(* IEC 61131-3 sources: iec-checker/test/st/bad, 2 files *)

(* ---- semantic-error.st ---- *)
TYPE
  ANALOG_DATA_OK: INT (0 .. 16);
  ANALOG_DATA_BAD: INT ("foo" .. "bar");
END_TYPE

(* ---- lexing-error.st ---- *)
PROGRAM program0
  VAR
    LocalVar0 : DINT;
    LocalVar1 : TOD;
    _LocalVar2 : DINT;
  END_VAR

  LocalVar0 := 42;

  wtf?
END_PROGRAM
